Universal Robots PolyScope program: TgtProg.urp

Program TgtProg (createdIn=3.0.0 lastSavedIn=3.0.0 directory=/programs installation=default)
Robot Program (runOnlyOnce=true motionType=MoveJ speed=1.047198 acceleration=1.396263 useActiveTCP=false)
  'Program generated by RoboDK v6.0.7 for UR10 on XX/XX/XXXX 18:00:00'
  'Using nominal kinematics.'
  Script: movej([0.174533, -0.174533, 0.349066, 0.000000, 0.523599, 0.000000],1.20000,0.75000,0,0.0000)
  Script: movej([0.174533, -0.174533, 0.349066, 0.000000, 0.523599, 0.000000],1.20000,0.75000,0,0.0000)
  Script: movej([0.174533, -0.174533, 0.349066, 0.000000, 0.523599, 0.000000],1.20000,0.75000,0,0.0000)
  Script: movej([0.174533, -0.174533, 0.349066, 0.000000, 0.523599, 0.000000],1.20000,0.75000,0,0.0000)
  Script: movej([0.174533, -0.174533, 0.349066, 0.000000, 0.523599, 0.000000],1.20000,0.75000,0,0.0000)
  Script: movej([0.174533, -0.174533, 0.349066, 0.000000, 0.523599, 0.000000],1.20000,0.75000,0,0.0000)
  Script: movej([0.174533, -0.174533, 0.349066, 0.000000, 0.523599, 0.000000],1.20000,0.75000,0,0.0000)
